Fanuc KAREL source: KO00090.KL

PROGRAM KO00090
%NOLOCKGROUP
%ENVIRONMENT MIR
VAR
  P1: JOINTPOS
  P2: XYZWPREXT
  F: BOOLEAN
  OUT: XYZWPR
BEGIN
  F = TRUE
  OUT = MIRROR(P1, P2, F)
END KO00090
